Staubli VAL3: insertCASE.pgx

public program insertCASE(string x_sKey, num x_nIndex, string x_sTRAJname, bool& x_bToSave, num x_nSwitchValue, num x_nType)
  local num l_nIndex
  local num l_i
begin

  if x_nIndex==0 and progTemp:pProgItem[x_sKey].pProgTemplate[x_nIndex].sTRAJname==""
    progTemp:pProgItem[x_sKey].pProgTemplate[x_nIndex].nType=6
    if x_nType==1
      progTemp:pProgItem[x_sKey].pProgTemplate[x_nIndex].sTRAJname="PROG"
    elseIf x_nType==2
      progTemp:pProgItem[x_sKey].pProgTemplate[x_nIndex].sTRAJname="TRAJ"
    endIf
    progTemp:pProgItem[x_sKey].pProgTemplate[x_nIndex].sSwitchItem.sIOValue=x_sTRAJname
    progTemp:pProgItem[x_sKey].pProgTemplate[x_nIndex].sSwitchItem.nSwitchValue=x_nSwitchValue
  else
    l_nIndex=x_nIndex+1
    //insert(progTemp:pProgItem[x_sKey].pProgTemplate[x_nIndex+1])
    append(progTemp:pProgItem[x_sKey].pProgTemplate)
    for l_i = size(progTemp:pProgItem[x_sKey].pProgTemplate)-1 to l_nIndex step -1
      call copyPara(x_sKey,l_i-1,l_i)
    endFor
    //insert(progTemp:pProgItem[x_sKey].pProgTemplate[x_nIndex+1])
    progTemp:pProgItem[x_sKey].pProgTemplate[x_nIndex+1].nType=6
    if x_nType==1
      progTemp:pProgItem[x_sKey].pProgTemplate[x_nIndex+1].sTRAJname="PROG"
    elseIf x_nType==2
      progTemp:pProgItem[x_sKey].pProgTemplate[x_nIndex+1].sTRAJname="TRAJ"
    endIf
    progTemp:pProgItem[x_sKey].pProgTemplate[x_nIndex+1].sSwitchItem.sIOValue=x_sTRAJname
    progTemp:pProgItem[x_sKey].pProgTemplate[x_nIndex+1].sSwitchItem.nSwitchValue=x_nSwitchValue
  endIf

  x_bToSave=true
end
